SUBAPPLICATION Dom (* Subapplication Type *)
  (* Standard: 61499-2 *)
  (* Version 1.0, 2023-01-29, Franz *)
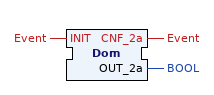
  EVENT_INPUT
    INIT;
  END_EVENT
  EVENT_OUTPUT
    CNF_2a;
  END_EVENT
  VAR_OUTPUT
    OUT_2a : BOOL;
  END_VAR
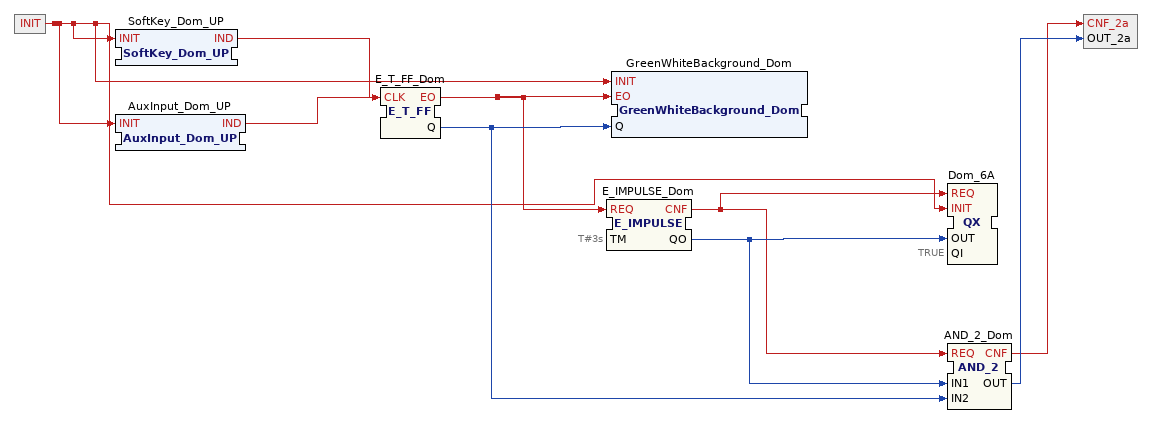
  FBS
    AND_2_Dom : AND_2;
    E_T_FF_Dom : E_T_FF;
    Dom_6A : QX(QI := TRUE);
    E_IMPULSE_Dom : E_IMPULSE(TM := T#3s);
  END_FBS
  SUBAPPS
    GreenWhiteBackground_Dom : GreenWhiteBackground_Dom;
    AuxInput_Dom_UP : AuxInput_Dom_UP;
    SoftKey_Dom_UP : SoftKey_Dom_UP;
  END_SUBAPPS
  EVENT_CONNECTIONS
    E_IMPULSE_Dom.CNF TO AND_2_Dom.REQ;
    E_T_FF_Dom.EO TO E_IMPULSE_Dom.REQ;
    E_IMPULSE_Dom.CNF TO Dom_6A.REQ;
    AND_2_Dom.CNF TO CNF_2a;
    INIT TO Dom_6A.INIT;
    INIT TO GreenWhiteBackground_Dom.INIT;
    E_T_FF_Dom.EO TO GreenWhiteBackground_Dom.EO;
    INIT TO AuxInput_Dom_UP.INIT;
    AuxInput_Dom_UP.IND TO E_T_FF_Dom.CLK;
    INIT TO SoftKey_Dom_UP.INIT;
    SoftKey_Dom_UP.IND TO E_T_FF_Dom.CLK;
  END_CONNECTIONS
  DATA_CONNECTIONS
    E_IMPULSE_Dom.QO TO AND_2_Dom.IN1;
    E_T_FF_Dom.Q TO AND_2_Dom.IN2; (* Schieber offen *)
    E_IMPULSE_Dom.QO TO Dom_6A.OUT;
    AND_2_Dom.OUT TO OUT_2a;
    E_T_FF_Dom.Q TO GreenWhiteBackground_Dom.Q; (* Schieber offen *)
  END_CONNECTIONS
END_SUBAPPLICATION
